TYPE st_LineSourceValves :
STRUCT
	valTankA				:	E_Pis_Name	;
	valTankB				:	E_Pis_Name	;
	valTapWater				:	E_Pis_Name	;
	valTapWater_esle		:	E_Pis_Name	;
	valTapWater_Drain		:	E_Pis_Name	;	
	valDrain				:	E_Pis_Name	;
	valCIP					:	E_Pis_Name	;
	valCIP_Sel				:	E_Pis_Name	;
	valBlockWater			:	E_Pis_Name	;	
	valWaterSource			:	E_Pis_Name	;
	valWaterSource_Drain	:	E_Pis_Name	;
END_STRUCT
END_TYPE

(* stored: Version 1.1.0.1, ProductVersion 3.1.4024.15
   DUT st_LineSourceValves: Id {a41f72ff-52c6-46d7-bb38-ed2f21ade05a} *)
